//{attribute 'qualified_only'}
VAR_GLOBAL
	ErrorAcknowledgement AT %Q*: BOOL;
	Run AT %Q*: BOOL;
	SEW_Safety_Reset	AT %Q*: BOOL;
END_VAR

(* stored: Version 1.1.0.1
   GVL IO_Safety: Id {9e5608f6-3ba4-46d2-a5f1-03831b3c3045} *)
